(* IEC 61131-3 sources: s7-to-codesys/tests/POUs/S7Compat/FB_StandardCounter_Test, 4 files *)

(* ---- CtdStopsAtZero.method.decl.st ---- *)
// CTD: LOAD по уровню ставит CV := PV, фронт CD уменьшает CV, но не ниже 0; Q = (CV = 0).
METHOD PRIVATE CtdStopsAtZero
VAR
    fbDut : CTD;    // проверяемый счётчик (новый экземпляр на каждый вызов метода)
END_VAR

(* ---- CtuCountsRisingEdges.method.decl.st ---- *)
// CTU: CV растёт только по фронту CU, Q = CV >= PV, RESET по уровню обнуляет CV.
METHOD PRIVATE CtuCountsRisingEdges
VAR
    fbDut : CTU;    // проверяемый счётчик (новый экземпляр на каждый вызов метода)
END_VAR

(* ---- CtudBothEdgesSameCall.method.decl.st ---- *)
// CTUD: фронты CU и CD в одном вызове — модель stsim применяет оба (+1 и -1), CV не меняется.
// Справка Standard этот случай не описывает; тест фиксирует поведение 3.5.17.0.
METHOD PRIVATE CtudBothEdgesSameCall
VAR
    fbDut : CTUD;   // проверяемый счётчик (новый экземпляр на каждый вызов метода)
END_VAR

(* ---- CtudResetBeatsLoad.method.decl.st ---- *)
// CTUD: RESET и LOAD одновременно — RESET главнее (CV = 0); QU = CV >= PV, QD = (CV = 0).
METHOD PRIVATE CtudResetBeatsLoad
VAR
    fbDut : CTUD;   // проверяемый счётчик (новый экземпляр на каждый вызов метода)
END_VAR
